// TIA Portal V20 export
// export: Created 2026-10-12T05:06:04.4259791Z, ExportSetting WithDefaults, DisplayName Totally Integrated Automation Portal, DisplayVersion V20, DisplayName TIA Portal Openness, DisplayVersion V20, DisplayName TIA Portal Teamcenter Gateway, DisplayVersion V20, DisplayName TIA Portal Version Control Interface, DisplayVersion V20, DisplayName SINAMICS Startdrive Advanced, DisplayVersion V20 SP1 Update 2, DisplayName SINAMICS Startdrive G110M, G120, G120C, G120D, G120P, G115D, DisplayVersion V20 SP1 Update 2, DisplayName SINAMICS Startdrive G130, G150, S120, S150, SINAMICS MV, G220, S200, S210, DisplayVersion V20 SP1 Update 2, DisplayName STEP 7 Professional, DisplayVersion V20, DisplayName STEP 7 Safety, DisplayVersion V20, DisplayName WinCC Basic/Comfort/Advanced, DisplayVersion V20, DisplayName WinCC Professional, DisplayVersion V20, DisplayName WinCC Unified, DisplayVersion V20
FUNCTION "FRK_ConfigDecode" : Bool   // FC95, SCL
{ S7_Optimized_Access := 'TRUE' }
VERSION : 0.1
// Keyed local-retain config. The typed owner validates before publishing a value.
// stored: AutoNumber true, IsIECCheckEnabled false, SetENOAutomatically false, UDAEnableTagReadback false
   VAR_INPUT
      Text : WString;
      Storage : DInt;
      Minimum : LReal;
      Maximum : LReal;
      MaxLength : Int;
   END_VAR
   VAR_IN_OUT
      Value : "FRK_ConfigValue";
   END_VAR
   VAR_TEMP
      Index : Int;
      Width : Int;
      Negative : Bool;
      Magnitude : ULInt;
      Digit : ULInt;
   END_VAR
BEGIN

   #FRK_ConfigDecode := FALSE;
   IF #Storage = 8 THEN
       IF LEN(#Text) > #MaxLength THEN
           RETURN;
       END_IF;
       #Value.Text := WSTRING_TO_STRING(#Text);
       IF STRING_TO_WSTRING(#Value.Text) <> #Text THEN
           RETURN;
       END_IF;
       #FRK_ConfigDecode := TRUE;
       RETURN;
   END_IF;
   IF #Storage = 1 THEN
       IF #Text = WSTRING#'true' OR #Text = WSTRING#'TRUE' OR #Text = WSTRING#'1' THEN
           #Value.Flag := TRUE;
       ELSIF #Text = WSTRING#'false' OR #Text = WSTRING#'FALSE' OR #Text = WSTRING#'0' THEN
           #Value.Flag := FALSE;
       ELSE
           RETURN;
       END_IF;
       #FRK_ConfigDecode := TRUE;
       RETURN;
   END_IF;
   #Width := LEN(#Text);
   IF #Width = 0 THEN
       RETURN;
   END_IF;
   #Negative := FALSE;
   #Index := 1;
   IF #Text[1] = WCHAR#'-' THEN
       #Negative := TRUE;
       #Index := 2;
   ELSIF #Text[1] = WCHAR#'+' THEN
       #Index := 2;
   END_IF;
   IF #Index > #Width THEN
       RETURN;
   END_IF;
   #Magnitude := 0;
   WHILE #Index <= #Width DO
       IF #Text[#Index] < WCHAR#'0' OR #Text[#Index] > WCHAR#'9' THEN
           RETURN;
       END_IF;
       #Digit := UINT_TO_ULINT(WCHAR_TO_UINT(#Text[#Index]) - UINT#48);
       IF #Magnitude > (ULINT#4294967295 - #Digit) / ULINT#10 THEN
           RETURN;
       END_IF;
       #Magnitude := #Magnitude * ULINT#10 + #Digit;
       #Index := #Index + 1;
   END_WHILE;
   #Value.Number := ULINT_TO_LINT(#Magnitude);
   IF #Negative THEN
       #Value.Number := - #Value.Number;
   END_IF;
   IF LINT_TO_LREAL(#Value.Number) < #Minimum OR LINT_TO_LREAL(#Value.Number) > #Maximum THEN
       RETURN;
   END_IF;
   #FRK_ConfigDecode := TRUE;
END_FUNCTION
